INTERFACE I_FixtureDevice

METHOD Reset : BOOL
VAR_INPUT
END_VAR
END_METHOD

END_INTERFACE

(* stored: Version 1.1.0.1
   Itf I_FixtureDevice: Id {c02bec33-8a03-40cd-be22-7cfa07d56327}
   Method Reset: Id {f72165a0-e4d0-4e8c-b08d-702c655ed0e0} *)
